(* IEC 61131-3 sources: RootPLC/conformance/cases/runtime, 8 files *)

(* ---- err_located_type_mismatch.st ---- *)
(* spec: [runtime.image.type]
   expect: error RP0205 *)
PROGRAM Mismatch
VAR
    level AT %IX0.0 : INT;
END_VAR
level := level + 1;
END_PROGRAM

(* ---- ok_deploy_warm_start.st ---- *)
(* spec: [runtime.deploy] [runtime.retain]
   expect: ok *)
(* Version 2 of a counter program, as it would be deployed over version 1:
   `total` (RETAIN, same name and type) keeps its value across the swap;
   `rate` is new and starts from its initial value. *)
PROGRAM Counter
VAR RETAIN
    total : UDINT;
END_VAR
VAR
    btn AT %IX0.0 : BOOL;
    edge : R_TRIG;
    rate : UINT := 1;
END_VAR
edge(CLK := btn);
IF edge.Q THEN
    total := total + UINT_TO_UDINT(rate);
END_IF;
END_PROGRAM

(* ---- ok_engine_c_io.st ---- *)
(* spec: [build.c.abi] [build.c.shim] [build.c.shim.services] [runtime.engine] [runtime.image] [runtime.retain]
   expect: ok *)
(* Located inputs, outputs and memory, a RETAIN counter and a timer:
   crates/rootplc-driver/tests/engine_c.rs runs this program on the VM
   engine, the C engine (rootplc runtime --engine c) and the C runtime
   (runtime-c, POSIX port) under the same virtual clock and inputs, and
   compares the variables and the output image. *)
PROGRAM PRG_Io
VAR
    start AT %IX0.0 : BOOL;
    level AT %IW2 : INT;
    lamp AT %QX0.1 : BOOL;
    speed AT %QW2 : INT;
    hold AT %MD4 : REAL;
    count : DINT;
    blink : TON;
    tally AT %QB4 : USINT;
END_VAR
VAR RETAIN
    starts : UDINT;
END_VAR
count := count + 1;
lamp := start AND NOT blink.Q;
blink(IN := start AND NOT blink.Q, PT := T#30ms);
IF blink.Q THEN
    starts := starts + 1;
END_IF;
speed := level * 2;
hold := INT_TO_REAL(level) / 3.0;
tally := DINT_TO_USINT(count);
END_PROGRAM

(* ---- ok_located_types.st ---- *)
(* spec: [runtime.image] [runtime.image.type] [variables.located]
   expect: ok *)
(* Every size letter with a type that fits it. *)
PROGRAM Located
VAR
    start_btn AT %IX0.0 : BOOL;
    stop_btn  AT %I0.1 : BOOL;
    level     AT %IW2 : INT;
    raw_byte  AT %IB4 : BYTE;
    flag_byte AT %IB5 : BOOL;
    count     AT %ID8 : UDINT;
    scale     AT %MD0 : REAL;
    total     AT %ML8 : LREAL;
    pump      AT %QX0.0 : BOOL;
    speed     AT %QW2 : UINT;
END_VAR
pump := start_btn AND NOT stop_btn;
speed := INT_TO_UINT(level);
total := total + REAL_TO_LREAL(scale);
END_PROGRAM

(* ---- ok_modbus_image.st ---- *)
(* spec: [runtime.modbus] [runtime.image]
   expect: ok *)
(* A program whose image an HMI reads and sets over Modbus TCP: the set
   point in %MW0 is holding register 0, the measured level %IW0 is input
   register 0, the pump output %QX0.0 is coil 0. *)
PROGRAM Tank
VAR
    setpoint AT %MW0 : INT;
    level    AT %IW0 : INT;
    pump     AT %QX0.0 : BOOL;
END_VAR
pump := level < setpoint;
END_PROGRAM

(* ---- ok_retain_section.st ---- *)
(* spec: [runtime.retain] [variables.section]
   expect: ok *)
(* Counters that survive a restart of the runtime: a RETAIN section of the
   program and of a global variable list. *)
CONFIGURATION Plant
    VAR_GLOBAL RETAIN
        hours : UDINT;
    END_VAR
    RESOURCE Cpu ON PLC
        TASK Main (INTERVAL := T#10ms, PRIORITY := 1);
        PROGRAM Run WITH Main : Counter;
    END_RESOURCE
END_CONFIGURATION

PROGRAM Counter
VAR_EXTERNAL
    hours : UDINT;
END_VAR
VAR RETAIN
    starts : UDINT;
END_VAR
VAR
    btn AT %IX0.0 : BOOL;
    edge : R_TRIG;
END_VAR
edge(CLK := btn);
IF edge.Q THEN
    starts := starts + 1;
END_IF;
END_PROGRAM

(* ---- ok_runtime_cycle_program.st ---- *)
(* spec: [runtime.cycle] [runtime.watchdog] [runtime.status]
   expect: ok
   run: Blink cycles=50 *)
(* A program as the runtime runs it: inputs and outputs are located, one
   call per cycle, time from the cycle clock. Under the runtime a fault in a
   cycle (here none) would stop it with safe outputs. *)
PROGRAM Blink
VAR
    lamp AT %QX0.0 : BOOL;
    t : TON;
    n : INT;
END_VAR
t(IN := NOT t.Q, PT := T#100ms);
IF t.Q THEN
    lamp := NOT lamp;
    n := n + 1;
END_IF;
END_PROGRAM

(* ---- warn_located_byte_offset.st ---- *)
(* spec: [runtime.image.type] [scope.vendor-forms]
   expect: warning RP0135 *)
(* The TwinCAT reading of a byte, word, double or long address: the number
   is the byte offset, the type gives the size (Beckhoff samples place REAL,
   LREAL and DINT at %MB addresses this way). *)
PROGRAM ByteOffset
VAR
    lamp  AT %QW0 : BOOL;
    level AT %MB20 : REAL;
    total AT %MB24 : LREAL;
    count AT %MB32 : DINT;
END_VAR
lamp := TRUE;
level := level + 0.5;
count := count + 1;
END_PROGRAM
